// TIA Portal V21 export
// export: Created 2026-10-12T11:32:16.8302894Z, ExportSetting WithDefaults, DisplayName Totally Integrated Automation Portal, DisplayVersion V21, DisplayName STEP 7 Professional, DisplayVersion V21, DisplayName STEP 7 Safety, DisplayVersion V21, DisplayName Tech WebApplication, DisplayVersion V21, DisplayName WinCC Basic/Comfort/Advanced, DisplayVersion V21, DisplayName WinCC Unified, DisplayVersion V21
FUNCTION "FC_TCP_IP" : Void   // FC6, LAD
{ S7_Optimized_Access := 'TRUE' }
VERSION : 0.1
// stored: AutoNumber true, IsIECCheckEnabled false, SetENOAutomatically false, UDAEnableTagReadback false
BEGIN

REGION Network 1: Connection definition
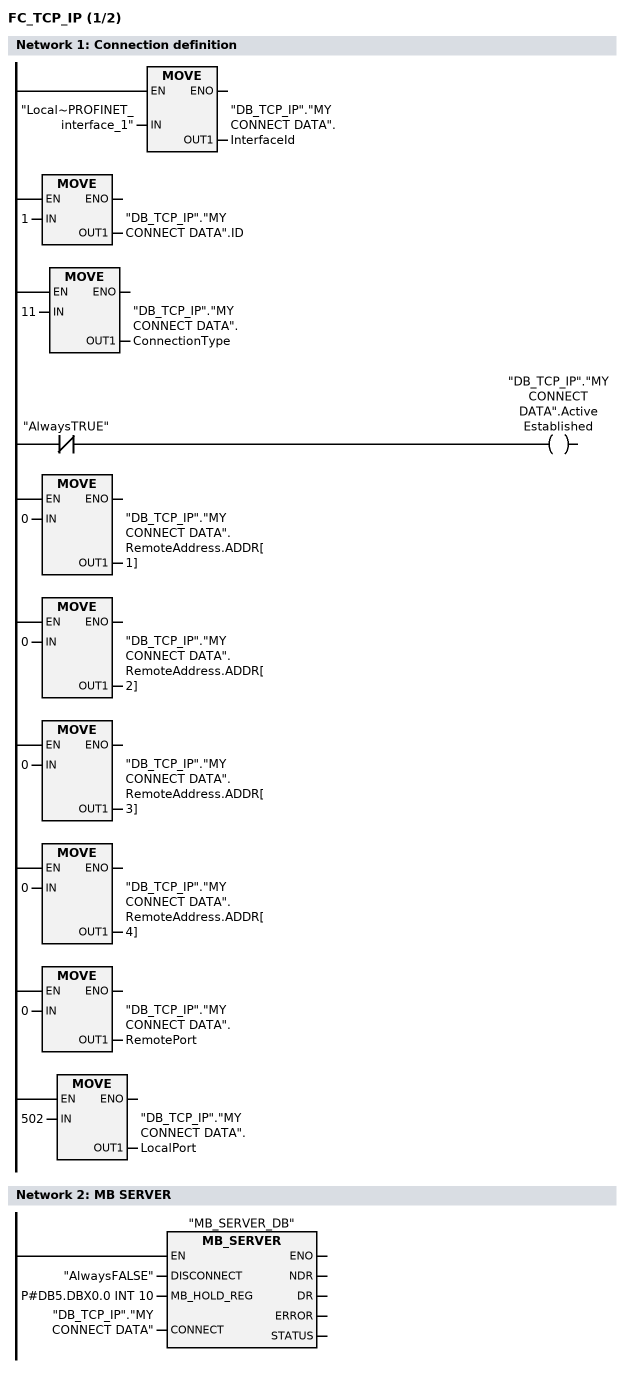
   RUNG wire#powerrail
      Move(in := "Local~PROFINET_interface_1", out1 => "DB_TCP_IP"."MY CONNECT DATA".InterfaceId)
   END_RUNG
   RUNG wire#powerrail
      Move(in := 1, out1 => "DB_TCP_IP"."MY CONNECT DATA".ID)
   END_RUNG
   RUNG wire#powerrail
      Move(in := 11, out1 => "DB_TCP_IP"."MY CONNECT DATA".ConnectionType)
   END_RUNG
   RUNG wire#powerrail
      I_Contact( "AlwaysTRUE" )
      Coil( "DB_TCP_IP"."MY CONNECT DATA".ActiveEstablished )
   END_RUNG
   RUNG wire#powerrail
      Move(in := 0, out1 => "DB_TCP_IP"."MY CONNECT DATA".RemoteAddress.ADDR[1])
   END_RUNG
   RUNG wire#powerrail
      Move(in := 0, out1 => "DB_TCP_IP"."MY CONNECT DATA".RemoteAddress.ADDR[2])
   END_RUNG
   RUNG wire#powerrail
      Move(in := 0, out1 => "DB_TCP_IP"."MY CONNECT DATA".RemoteAddress.ADDR[3])
   END_RUNG
   RUNG wire#powerrail
      Move(in := 0, out1 => "DB_TCP_IP"."MY CONNECT DATA".RemoteAddress.ADDR[4])
   END_RUNG
   RUNG wire#powerrail
      Move(in := 0, out1 => "DB_TCP_IP"."MY CONNECT DATA".RemotePort)
   END_RUNG
   RUNG wire#powerrail
      Move(in := 502, out1 => "DB_TCP_IP"."MY CONNECT DATA".LocalPort)
   END_RUNG
   // the same network as SCL:
   "DB_TCP_IP"."MY CONNECT DATA".InterfaceId := "Local~PROFINET_interface_1";
   "DB_TCP_IP"."MY CONNECT DATA".ID := 1;
   "DB_TCP_IP"."MY CONNECT DATA".ConnectionType := 11;
   "DB_TCP_IP"."MY CONNECT DATA".ActiveEstablished := NOT "AlwaysTRUE";
   "DB_TCP_IP"."MY CONNECT DATA".RemoteAddress.ADDR[1] := 0;
   "DB_TCP_IP"."MY CONNECT DATA".RemoteAddress.ADDR[2] := 0;
   "DB_TCP_IP"."MY CONNECT DATA".RemoteAddress.ADDR[3] := 0;
   "DB_TCP_IP"."MY CONNECT DATA".RemoteAddress.ADDR[4] := 0;
   "DB_TCP_IP"."MY CONNECT DATA".RemotePort := 0;
   "DB_TCP_IP"."MY CONNECT DATA".LocalPort := 502;
END_REGION

REGION Network 2: MB SERVER
   RUNG wire#powerrail
      "MB_SERVER_DB".MB_SERVER(DISCONNECT := "AlwaysFALSE", MB_HOLD_REG := P#DB5.DBX0.0 INT 10, CONNECT := "DB_TCP_IP"."MY CONNECT DATA", NDR =>, DR =>, ERROR =>, STATUS =>)
   END_RUNG
   // the same network as SCL:
   "MB_SERVER_DB"(DISCONNECT := "AlwaysFALSE",   // MB_SERVER
                  MB_HOLD_REG := P#DB5.DBX0.0 INT 10,
                  CONNECT := "DB_TCP_IP"."MY CONNECT DATA");
END_REGION

REGION Network 3: ERROR CHECK
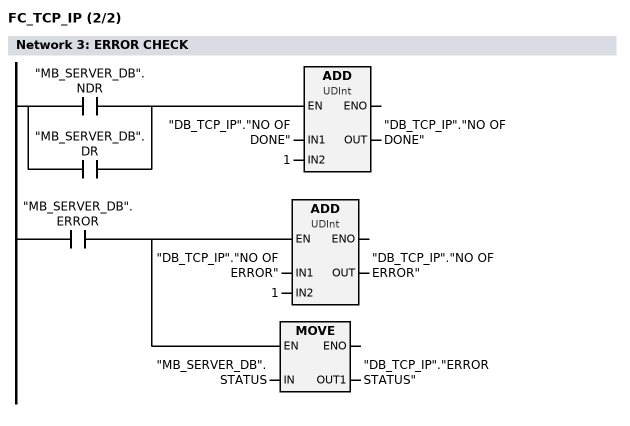
   RUNG wire#powerrail
      Contact( "MB_SERVER_DB".NDR )
      wire#w1
      { S7_Templates := "SrcType := UDInt" } Add(in1 := "DB_TCP_IP"."NO OF DONE", in2 := 1, out => "DB_TCP_IP"."NO OF DONE")
   END_RUNG
   RUNG wire#powerrail
      Contact( "MB_SERVER_DB".DR )
   END_RUNG wire#w1
   RUNG wire#powerrail
      Contact( "MB_SERVER_DB".ERROR )
      wire#w2
      { S7_Templates := "SrcType := UDInt" } Add(in1 := "DB_TCP_IP"."NO OF ERROR", in2 := 1, out => "DB_TCP_IP"."NO OF ERROR")
   END_RUNG
   RUNG wire#w2
      Move(in := "MB_SERVER_DB".STATUS, out1 => "DB_TCP_IP"."ERROR STATUS")
   END_RUNG
   // the same network as SCL:
   IF "MB_SERVER_DB".NDR OR "MB_SERVER_DB".DR THEN
       "DB_TCP_IP"."NO OF DONE" := "DB_TCP_IP"."NO OF DONE" + 1;
   END_IF;
   IF "MB_SERVER_DB".ERROR THEN
       "DB_TCP_IP"."NO OF ERROR" := "DB_TCP_IP"."NO OF ERROR" + 1;
       "DB_TCP_IP"."ERROR STATUS" := "MB_SERVER_DB".STATUS;
   END_IF;
END_REGION
END_FUNCTION
